// TIA Portal V21 export
// export: Created 2026-11-08T21:35:45.895519Z, ExportSetting WithDefaults, DisplayName Totally Integrated Automation Portal, DisplayVersion V21 Update 3, DisplayName STEP 7 Professional, DisplayVersion V21 Update 3, DisplayName STEP 7 Safety, DisplayVersion V21, DisplayName Tech WebApplication, DisplayVersion V21, DisplayName WinCC Basic/Comfort/Advanced, DisplayVersion V21 Update 3, DisplayName WinCC Unified, DisplayVersion V21 Update 3
FUNCTION_BLOCK "FB_StlC_060"   // FB85, STL
TITLE = STL call VARIANT_TO_DB_ANY
{ S7_Optimized_Access := 'TRUE' }
VERSION : 0.1
// stored: AutoNumber true, IsRetainMemResEnabled false, MemoryReserve 100, UDAEnableTagReadback false
   VAR_OUTPUT
      io : Int;
   END_VAR
   VAR_IN_OUT
      v : Variant;
   END_VAR
   VAR_TEMP
      dba : DB_ANY;
   END_VAR
BEGIN

NETWORK
TITLE = 060 VARIANT_TO_DB_ANY
      CALL  VARIANT_TO_DB_ANY
      ( in      := #v,
        Ret_Val := #dba,
        err     := #io
      );

NETWORK
TITLE = 061 DB_ANY_TO_VARIANT
      CALL  DB_ANY_TO_VARIANT
      ( in      := #dba,
        Ret_Val := #v,
        err     := #io
      );
END_FUNCTION_BLOCK
